// Mitsubishi GX Works2 project: B_v6_ladder   PLC: Q03UDE

PROGRAM MAIN
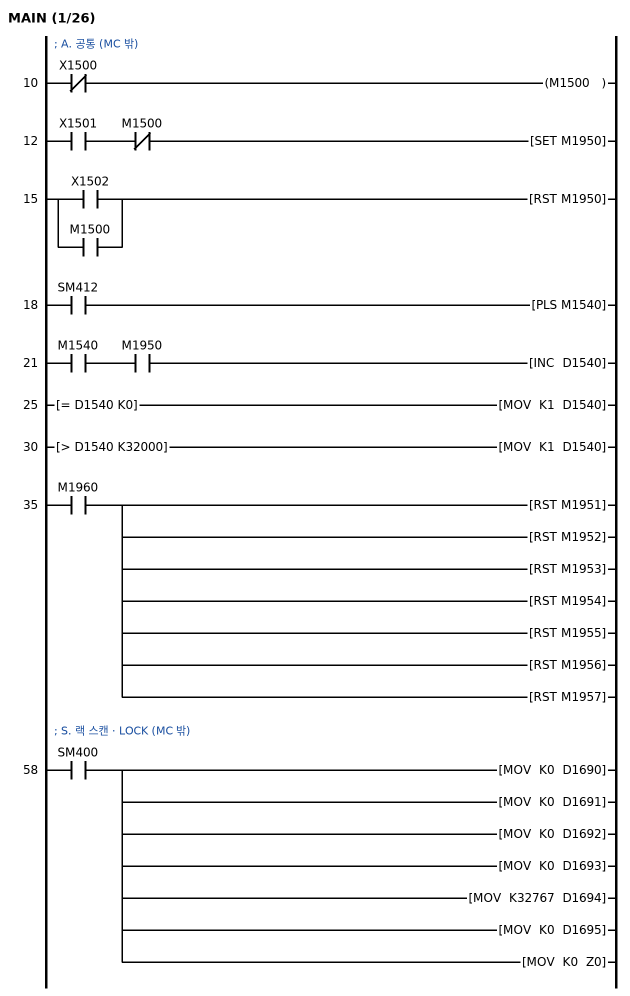
; A. 공통 (MC 밖)
10    LDI     X1500
      OUT     M1500
12    LD      X1501
      ANI     M1500
      SET     M1950
15    LD      X1502
      OR      M1500
      RST     M1950
18    LD      SM412
      PLS     M1540
21    LD      M1540
      AND     M1950
      INC     D1540
25    LD=     D1540 K0
      MOV     K1 D1540
30    LD>     D1540 K32000
      MOV     K1 D1540
35    LD      M1960
      RST     M1951
      RST     M1952
      RST     M1953
      RST     M1954
      RST     M1955
      RST     M1956
      RST     M1957
; S. 랙 스캔 · LOCK (MC 밖)
58    LD      SM400
      MOV     K0 D1690
      MOV     K0 D1691
      MOV     K0 D1692
      MOV     K0 D1693
      MOV     K32767 D1694
      MOV     K0 D1695
      MOV     K0 Z0
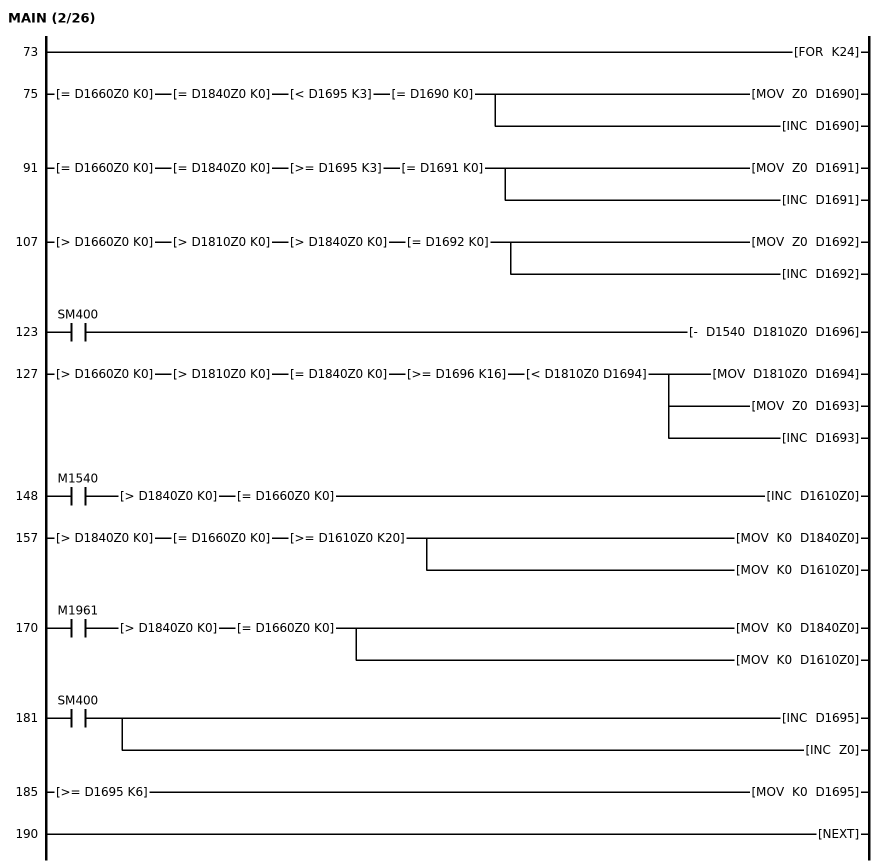
73    FOR     K24
75    LD=     D1660Z0 K0
      AND=    D1840Z0 K0
      AND<    D1695 K3
      AND=    D1690 K0
      MOV     Z0 D1690
      INC     D1690
91    LD=     D1660Z0 K0
      AND=    D1840Z0 K0
      AND>=   D1695 K3
      AND=    D1691 K0
      MOV     Z0 D1691
      INC     D1691
107   LD>     D1660Z0 K0
      AND>    D1810Z0 K0
      AND>    D1840Z0 K0
      AND=    D1692 K0
      MOV     Z0 D1692
      INC     D1692
123   LD      SM400
      -       D1540 D1810Z0 D1696
127   LD>     D1660Z0 K0
      AND>    D1810Z0 K0
      AND=    D1840Z0 K0
      AND>=   D1696 K16
      AND<    D1810Z0 D1694
      MOV     D1810Z0 D1694
      MOV     Z0 D1693
      INC     D1693
148   LD      M1540
      AND>    D1840Z0 K0
      AND=    D1660Z0 K0
      INC     D1610Z0
157   LD>     D1840Z0 K0
      AND=    D1660Z0 K0
      AND>=   D1610Z0 K20
      MOV     K0 D1840Z0
      MOV     K0 D1610Z0
170   LD      M1961
      AND>    D1840Z0 K0
      AND=    D1660Z0 K0
      MOV     K0 D1840Z0
      MOV     K0 D1610Z0
181   LD      SM400
      INC     D1695
      INC     Z0
185   LD>=    D1695 K6
      MOV     K0 D1695
190   NEXT
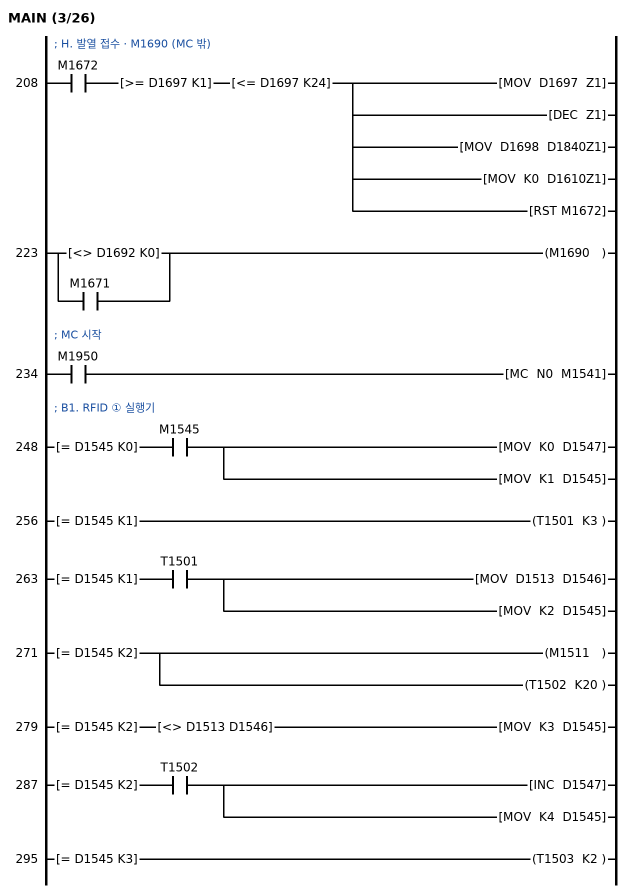
; H. 발열 접수 · M1690 (MC 밖)
208   LD      M1672
      AND>=   D1697 K1
      AND<=   D1697 K24
      MOV     D1697 Z1
      DEC     Z1
      MOV     D1698 D1840Z1
      MOV     K0 D1610Z1
      RST     M1672
223   LD<>    D1692 K0
      OR      M1671
      OUT     M1690
; MC 시작
234   LD      M1950
      MC      N0 M1541
; B1. RFID ① 실행기
248   LD=     D1545 K0
      AND     M1545
      MOV     K0 D1547
      MOV     K1 D1545
256   LD=     D1545 K1
      OUT     T1501 K3
263   LD=     D1545 K1
      AND     T1501
      MOV     D1513 D1546
      MOV     K2 D1545
271   LD=     D1545 K2
      OUT     M1511
      OUT     T1502 K20
279   LD=     D1545 K2
      AND<>   D1513 D1546
      MOV     K3 D1545
287   LD=     D1545 K2
      AND     T1502
      INC     D1547
      MOV     K4 D1545
295   LD=     D1545 K3
      OUT     T1503 K2
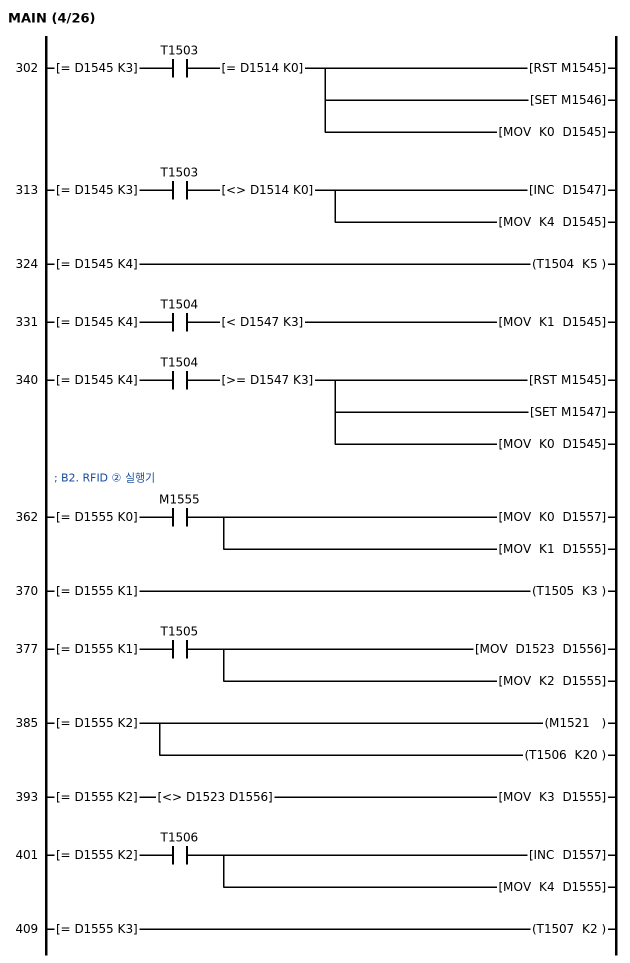
302   LD=     D1545 K3
      AND     T1503
      AND=    D1514 K0
      RST     M1545
      SET     M1546
      MOV     K0 D1545
313   LD=     D1545 K3
      AND     T1503
      AND<>   D1514 K0
      INC     D1547
      MOV     K4 D1545
324   LD=     D1545 K4
      OUT     T1504 K5
331   LD=     D1545 K4
      AND     T1504
      AND<    D1547 K3
      MOV     K1 D1545
340   LD=     D1545 K4
      AND     T1504
      AND>=   D1547 K3
      RST     M1545
      SET     M1547
      MOV     K0 D1545
; B2. RFID ② 실행기
362   LD=     D1555 K0
      AND     M1555
      MOV     K0 D1557
      MOV     K1 D1555
370   LD=     D1555 K1
      OUT     T1505 K3
377   LD=     D1555 K1
      AND     T1505
      MOV     D1523 D1556
      MOV     K2 D1555
385   LD=     D1555 K2
      OUT     M1521
      OUT     T1506 K20
393   LD=     D1555 K2
      AND<>   D1523 D1556
      MOV     K3 D1555
401   LD=     D1555 K2
      AND     T1506
      INC     D1557
      MOV     K4 D1555
409   LD=     D1555 K3
      OUT     T1507 K2
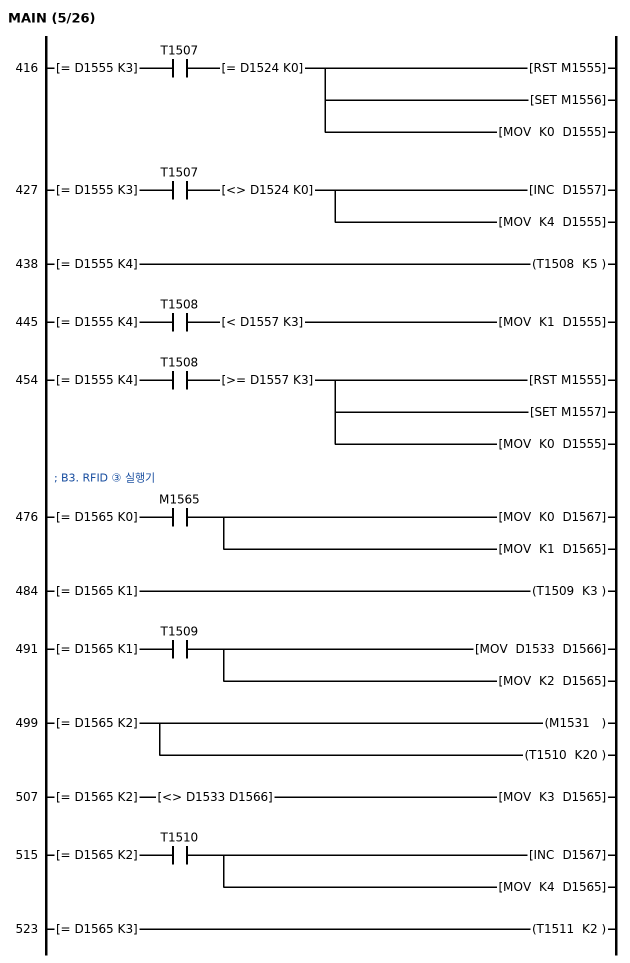
416   LD=     D1555 K3
      AND     T1507
      AND=    D1524 K0
      RST     M1555
      SET     M1556
      MOV     K0 D1555
427   LD=     D1555 K3
      AND     T1507
      AND<>   D1524 K0
      INC     D1557
      MOV     K4 D1555
438   LD=     D1555 K4
      OUT     T1508 K5
445   LD=     D1555 K4
      AND     T1508
      AND<    D1557 K3
      MOV     K1 D1555
454   LD=     D1555 K4
      AND     T1508
      AND>=   D1557 K3
      RST     M1555
      SET     M1557
      MOV     K0 D1555
; B3. RFID ③ 실행기
476   LD=     D1565 K0
      AND     M1565
      MOV     K0 D1567
      MOV     K1 D1565
484   LD=     D1565 K1
      OUT     T1509 K3
491   LD=     D1565 K1
      AND     T1509
      MOV     D1533 D1566
      MOV     K2 D1565
499   LD=     D1565 K2
      OUT     M1531
      OUT     T1510 K20
507   LD=     D1565 K2
      AND<>   D1533 D1566
      MOV     K3 D1565
515   LD=     D1565 K2
      AND     T1510
      INC     D1567
      MOV     K4 D1565
523   LD=     D1565 K3
      OUT     T1511 K2
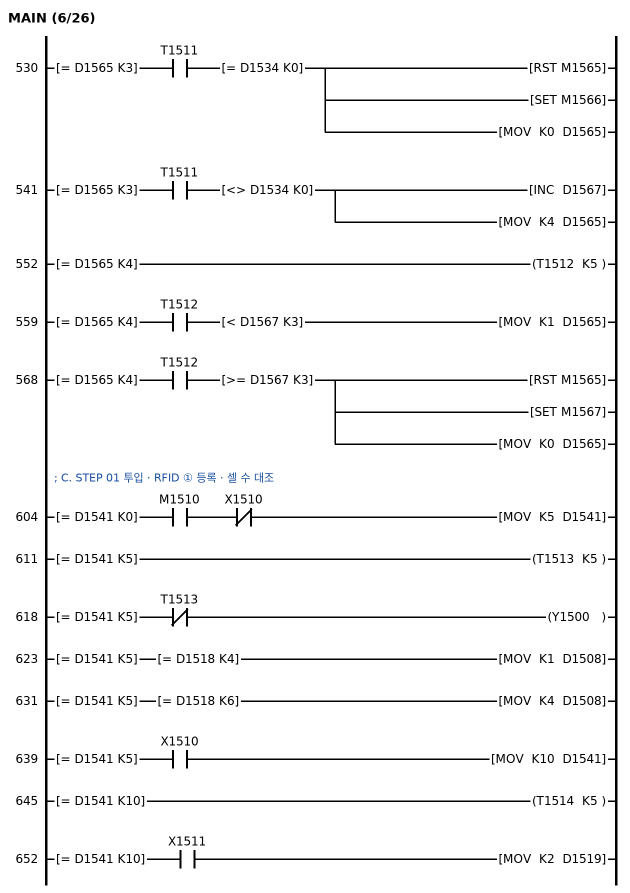
530   LD=     D1565 K3
      AND     T1511
      AND=    D1534 K0
      RST     M1565
      SET     M1566
      MOV     K0 D1565
541   LD=     D1565 K3
      AND     T1511
      AND<>   D1534 K0
      INC     D1567
      MOV     K4 D1565
552   LD=     D1565 K4
      OUT     T1512 K5
559   LD=     D1565 K4
      AND     T1512
      AND<    D1567 K3
      MOV     K1 D1565
568   LD=     D1565 K4
      AND     T1512
      AND>=   D1567 K3
      RST     M1565
      SET     M1567
      MOV     K0 D1565
; C. STEP 01 투입 · RFID ① 등록 · 셀 수 대조
604   LD=     D1541 K0
      AND     M1510
      ANI     X1510
      MOV     K5 D1541
611   LD=     D1541 K5
      OUT     T1513 K5
618   LD=     D1541 K5
      ANI     T1513
      OUT     Y1500
623   LD=     D1541 K5
      AND=    D1518 K4
      MOV     K1 D1508
631   LD=     D1541 K5
      AND=    D1518 K6
      MOV     K4 D1508
639   LD=     D1541 K5
      AND     X1510
      MOV     K10 D1541
645   LD=     D1541 K10
      OUT     T1514 K5
652   LD=     D1541 K10
      AND     X1511
      MOV     K2 D1519
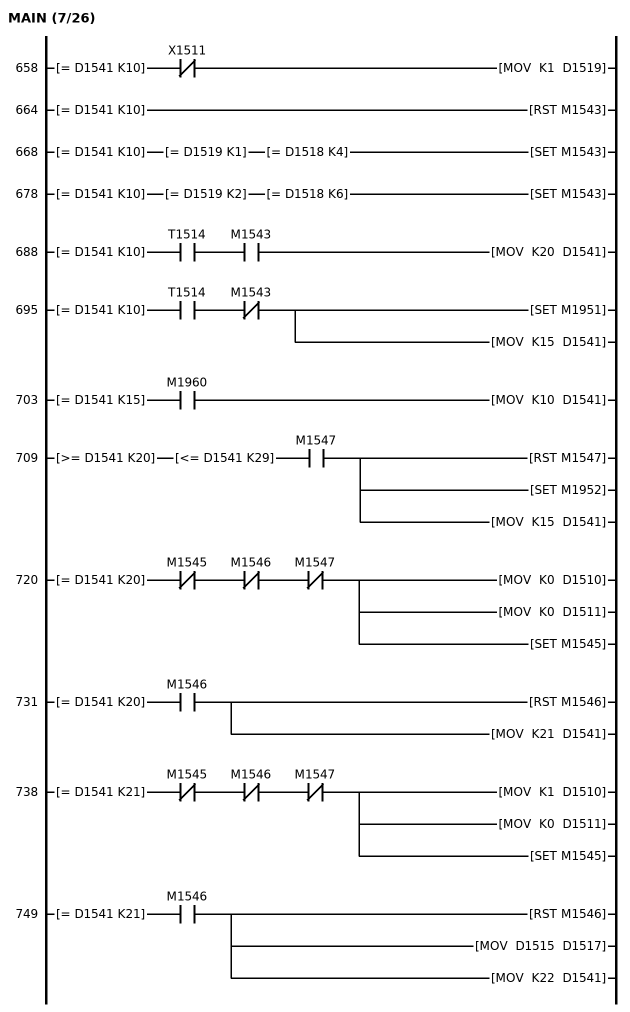
658   LD=     D1541 K10
      ANI     X1511
      MOV     K1 D1519
664   LD=     D1541 K10
      RST     M1543
668   LD=     D1541 K10
      AND=    D1519 K1
      AND=    D1518 K4
      SET     M1543
678   LD=     D1541 K10
      AND=    D1519 K2
      AND=    D1518 K6
      SET     M1543
688   LD=     D1541 K10
      AND     T1514
      AND     M1543
      MOV     K20 D1541
695   LD=     D1541 K10
      AND     T1514
      ANI     M1543
      SET     M1951
      MOV     K15 D1541
703   LD=     D1541 K15
      AND     M1960
      MOV     K10 D1541
709   LD>=    D1541 K20
      AND<=   D1541 K29
      AND     M1547
      RST     M1547
      SET     M1952
      MOV     K15 D1541
720   LD=     D1541 K20
      ANI     M1545
      ANI     M1546
      ANI     M1547
      MOV     K0 D1510
      MOV     K0 D1511
      SET     M1545
731   LD=     D1541 K20
      AND     M1546
      RST     M1546
      MOV     K21 D1541
738   LD=     D1541 K21
      ANI     M1545
      ANI     M1546
      ANI     M1547
      MOV     K1 D1510
      MOV     K0 D1511
      SET     M1545
749   LD=     D1541 K21
      AND     M1546
      RST     M1546
      MOV     D1515 D1517
      MOV     K22 D1541
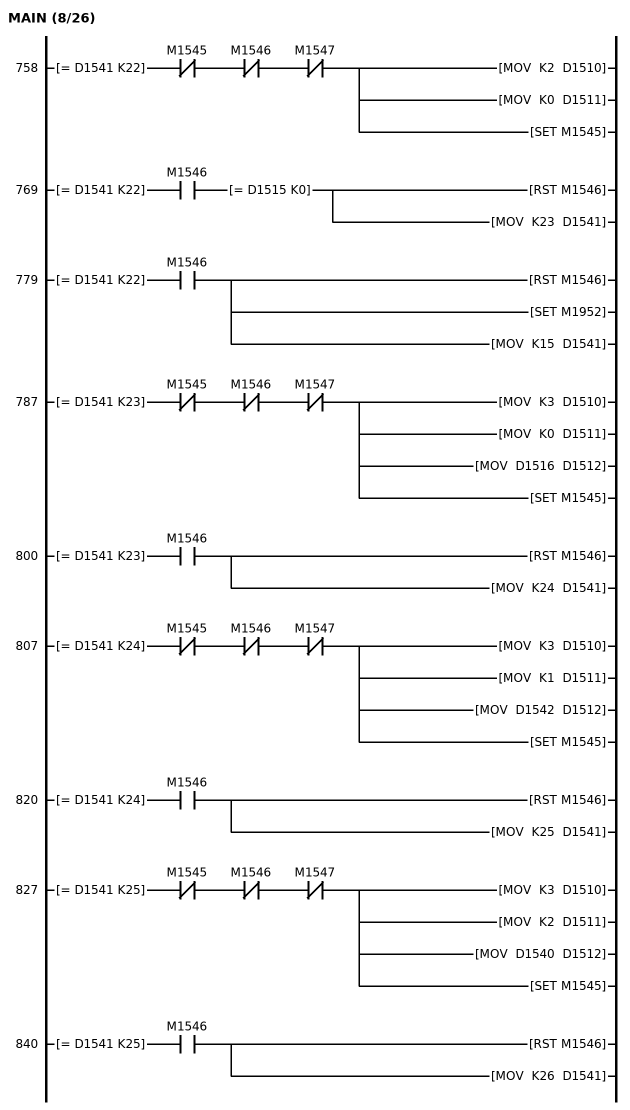
758   LD=     D1541 K22
      ANI     M1545
      ANI     M1546
      ANI     M1547
      MOV     K2 D1510
      MOV     K0 D1511
      SET     M1545
769   LD=     D1541 K22
      AND     M1546
      AND=    D1515 K0
      RST     M1546
      MOV     K23 D1541
779   LD=     D1541 K22
      AND     M1546
      RST     M1546
      SET     M1952
      MOV     K15 D1541
787   LD=     D1541 K23
      ANI     M1545
      ANI     M1546
      ANI     M1547
      MOV     K3 D1510
      MOV     K0 D1511
      MOV     D1516 D1512
      SET     M1545
800   LD=     D1541 K23
      AND     M1546
      RST     M1546
      MOV     K24 D1541
807   LD=     D1541 K24
      ANI     M1545
      ANI     M1546
      ANI     M1547
      MOV     K3 D1510
      MOV     K1 D1511
      MOV     D1542 D1512
      SET     M1545
820   LD=     D1541 K24
      AND     M1546
      RST     M1546
      MOV     K25 D1541
827   LD=     D1541 K25
      ANI     M1545
      ANI     M1546
      ANI     M1547
      MOV     K3 D1510
      MOV     K2 D1511
      MOV     D1540 D1512
      SET     M1545
840   LD=     D1541 K25
      AND     M1546
      RST     M1546
      MOV     K26 D1541
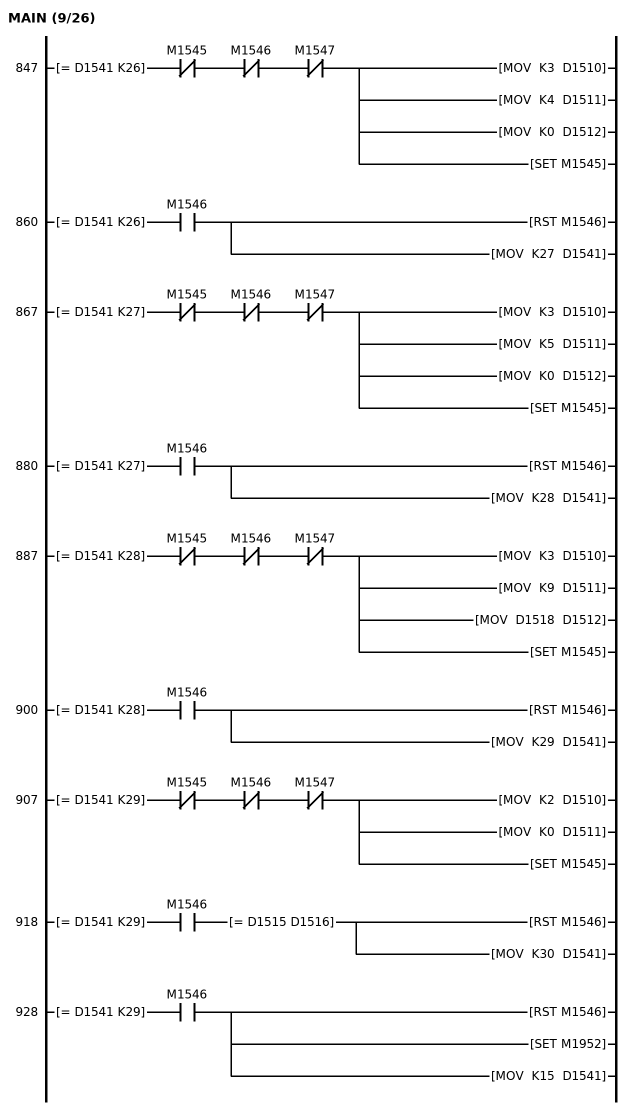
847   LD=     D1541 K26
      ANI     M1545
      ANI     M1546
      ANI     M1547
      MOV     K3 D1510
      MOV     K4 D1511
      MOV     K0 D1512
      SET     M1545
860   LD=     D1541 K26
      AND     M1546
      RST     M1546
      MOV     K27 D1541
867   LD=     D1541 K27
      ANI     M1545
      ANI     M1546
      ANI     M1547
      MOV     K3 D1510
      MOV     K5 D1511
      MOV     K0 D1512
      SET     M1545
880   LD=     D1541 K27
      AND     M1546
      RST     M1546
      MOV     K28 D1541
887   LD=     D1541 K28
      ANI     M1545
      ANI     M1546
      ANI     M1547
      MOV     K3 D1510
      MOV     K9 D1511
      MOV     D1518 D1512
      SET     M1545
900   LD=     D1541 K28
      AND     M1546
      RST     M1546
      MOV     K29 D1541
907   LD=     D1541 K29
      ANI     M1545
      ANI     M1546
      ANI     M1547
      MOV     K2 D1510
      MOV     K0 D1511
      SET     M1545
918   LD=     D1541 K29
      AND     M1546
      AND=    D1515 D1516
      RST     M1546
      MOV     K30 D1541
928   LD=     D1541 K29
      AND     M1546
      RST     M1546
      SET     M1952
      MOV     K15 D1541
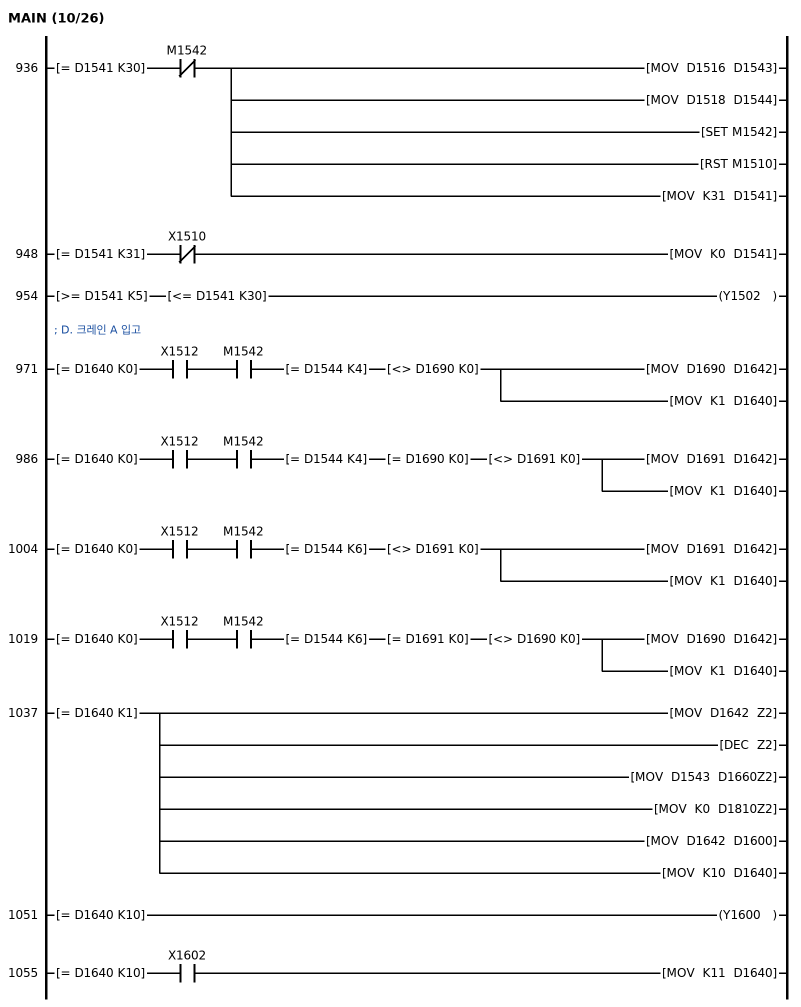
936   LD=     D1541 K30
      ANI     M1542
      MOV     D1516 D1543
      MOV     D1518 D1544
      SET     M1542
      RST     M1510
      MOV     K31 D1541
948   LD=     D1541 K31
      ANI     X1510
      MOV     K0 D1541
954   LD>=    D1541 K5
      AND<=   D1541 K30
      OUT     Y1502
; D. 크레인 A 입고
971   LD=     D1640 K0
      AND     X1512
      AND     M1542
      AND=    D1544 K4
      AND<>   D1690 K0
      MOV     D1690 D1642
      MOV     K1 D1640
986   LD=     D1640 K0
      AND     X1512
      AND     M1542
      AND=    D1544 K4
      AND=    D1690 K0
      AND<>   D1691 K0
      MOV     D1691 D1642
      MOV     K1 D1640
1004  LD=     D1640 K0
      AND     X1512
      AND     M1542
      AND=    D1544 K6
      AND<>   D1691 K0
      MOV     D1691 D1642
      MOV     K1 D1640
1019  LD=     D1640 K0
      AND     X1512
      AND     M1542
      AND=    D1544 K6
      AND=    D1691 K0
      AND<>   D1690 K0
      MOV     D1690 D1642
      MOV     K1 D1640
1037  LD=     D1640 K1
      MOV     D1642 Z2
      DEC     Z2
      MOV     D1543 D1660Z2
      MOV     K0 D1810Z2
      MOV     D1642 D1600
      MOV     K10 D1640
1051  LD=     D1640 K10
      OUT     Y1600
1055  LD=     D1640 K10
      AND     X1602
      MOV     K11 D1640
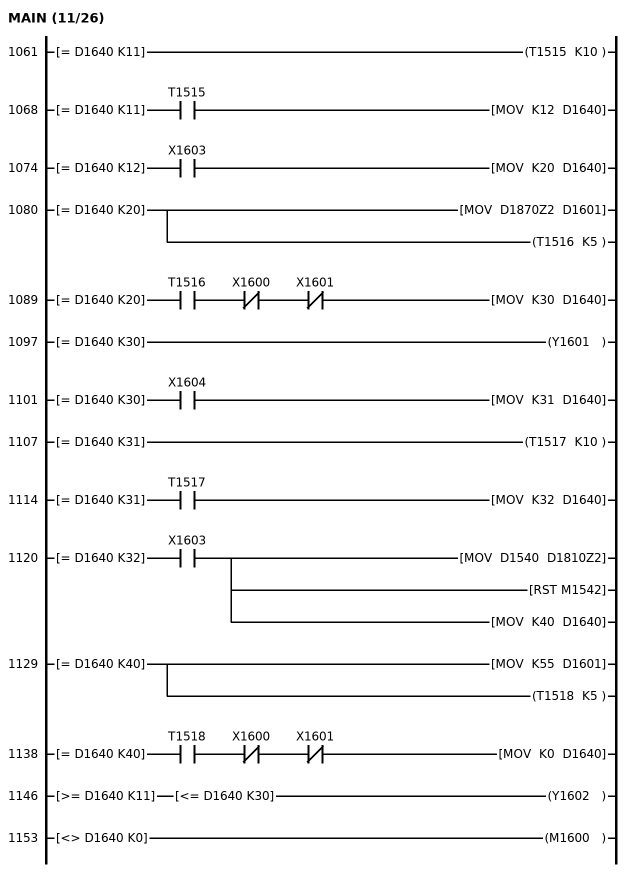
1061  LD=     D1640 K11
      OUT     T1515 K10
1068  LD=     D1640 K11
      AND     T1515
      MOV     K12 D1640
1074  LD=     D1640 K12
      AND     X1603
      MOV     K20 D1640
1080  LD=     D1640 K20
      MOV     D1870Z2 D1601
      OUT     T1516 K5
1089  LD=     D1640 K20
      AND     T1516
      ANI     X1600
      ANI     X1601
      MOV     K30 D1640
1097  LD=     D1640 K30
      OUT     Y1601
1101  LD=     D1640 K30
      AND     X1604
      MOV     K31 D1640
1107  LD=     D1640 K31
      OUT     T1517 K10
1114  LD=     D1640 K31
      AND     T1517
      MOV     K32 D1640
1120  LD=     D1640 K32
      AND     X1603
      MOV     D1540 D1810Z2
      RST     M1542
      MOV     K40 D1640
1129  LD=     D1640 K40
      MOV     K55 D1601
      OUT     T1518 K5
1138  LD=     D1640 K40
      AND     T1518
      ANI     X1600
      ANI     X1601
      MOV     K0 D1640
1146  LD>=    D1640 K11
      AND<=   D1640 K30
      OUT     Y1602
1153  LD<>    D1640 K0
      OUT     M1600
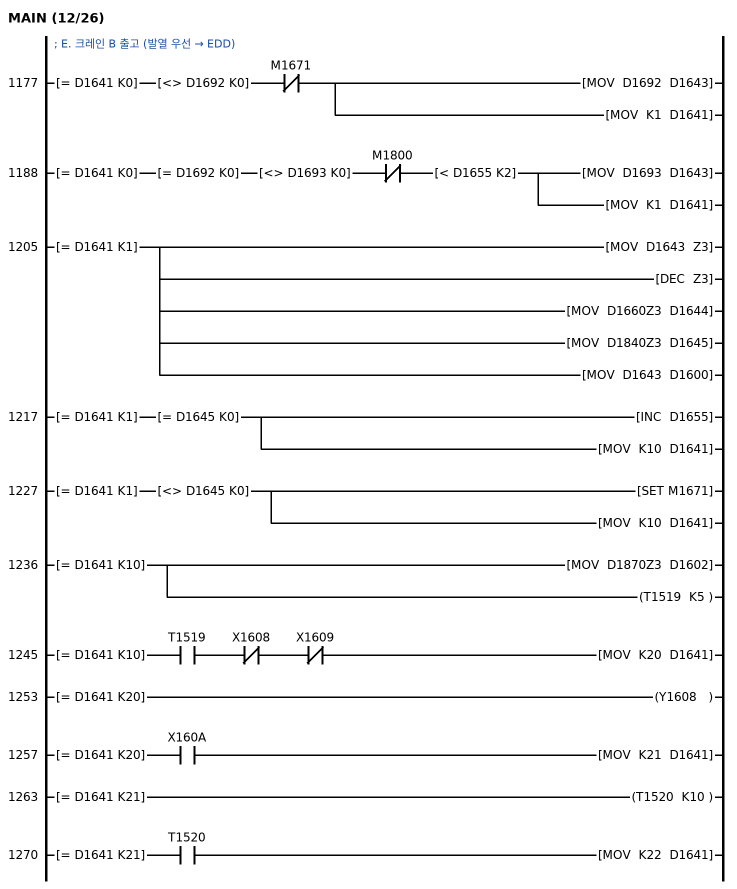
; E. 크레인 B 출고 (발열 우선 → EDD)
1177  LD=     D1641 K0
      AND<>   D1692 K0
      ANI     M1671
      MOV     D1692 D1643
      MOV     K1 D1641
1188  LD=     D1641 K0
      AND=    D1692 K0
      AND<>   D1693 K0
      ANI     M1800
      AND<    D1655 K2
      MOV     D1693 D1643
      MOV     K1 D1641
1205  LD=     D1641 K1
      MOV     D1643 Z3
      DEC     Z3
      MOV     D1660Z3 D1644
      MOV     D1840Z3 D1645
      MOV     D1643 D1600
1217  LD=     D1641 K1
      AND=    D1645 K0
      INC     D1655
      MOV     K10 D1641
1227  LD=     D1641 K1
      AND<>   D1645 K0
      SET     M1671
      MOV     K10 D1641
1236  LD=     D1641 K10
      MOV     D1870Z3 D1602
      OUT     T1519 K5
1245  LD=     D1641 K10
      AND     T1519
      ANI     X1608
      ANI     X1609
      MOV     K20 D1641
1253  LD=     D1641 K20
      OUT     Y1608
1257  LD=     D1641 K20
      AND     X160A
      MOV     K21 D1641
1263  LD=     D1641 K21
      OUT     T1520 K10
1270  LD=     D1641 K21
      AND     T1520
      MOV     K22 D1641
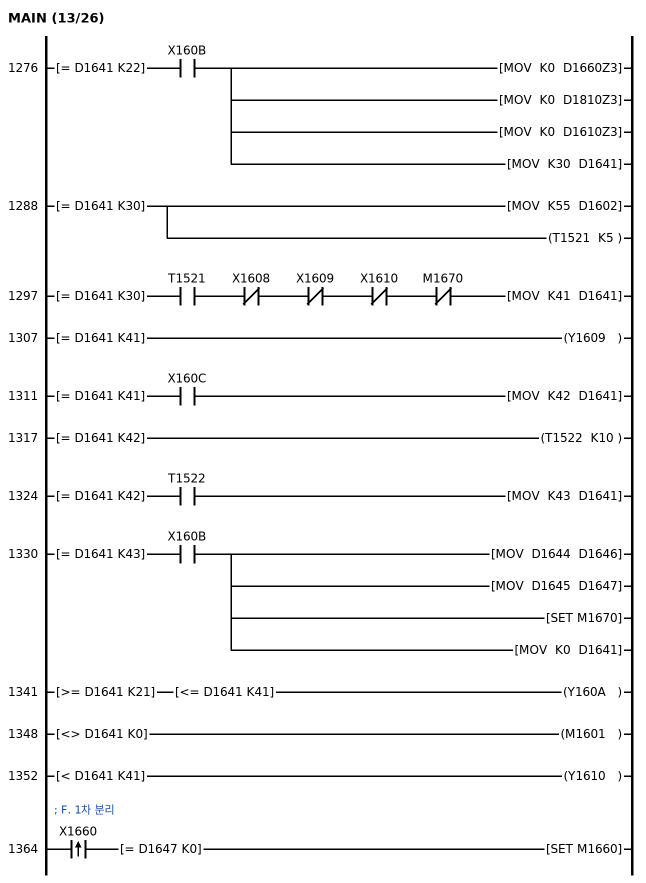
1276  LD=     D1641 K22
      AND     X160B
      MOV     K0 D1660Z3
      MOV     K0 D1810Z3
      MOV     K0 D1610Z3
      MOV     K30 D1641
1288  LD=     D1641 K30
      MOV     K55 D1602
      OUT     T1521 K5
1297  LD=     D1641 K30
      AND     T1521
      ANI     X1608
      ANI     X1609
      ANI     X1610
      ANI     M1670
      MOV     K41 D1641
1307  LD=     D1641 K41
      OUT     Y1609
1311  LD=     D1641 K41
      AND     X160C
      MOV     K42 D1641
1317  LD=     D1641 K42
      OUT     T1522 K10
1324  LD=     D1641 K42
      AND     T1522
      MOV     K43 D1641
1330  LD=     D1641 K43
      AND     X160B
      MOV     D1644 D1646
      MOV     D1645 D1647
      SET     M1670
      MOV     K0 D1641
1341  LD>=    D1641 K21
      AND<=   D1641 K41
      OUT     Y160A
1348  LD<>    D1641 K0
      OUT     M1601
1352  LD<     D1641 K41
      OUT     Y1610
; F. 1차 분리
1364  LDP     X1660
      AND=    D1647 K0
      SET     M1660
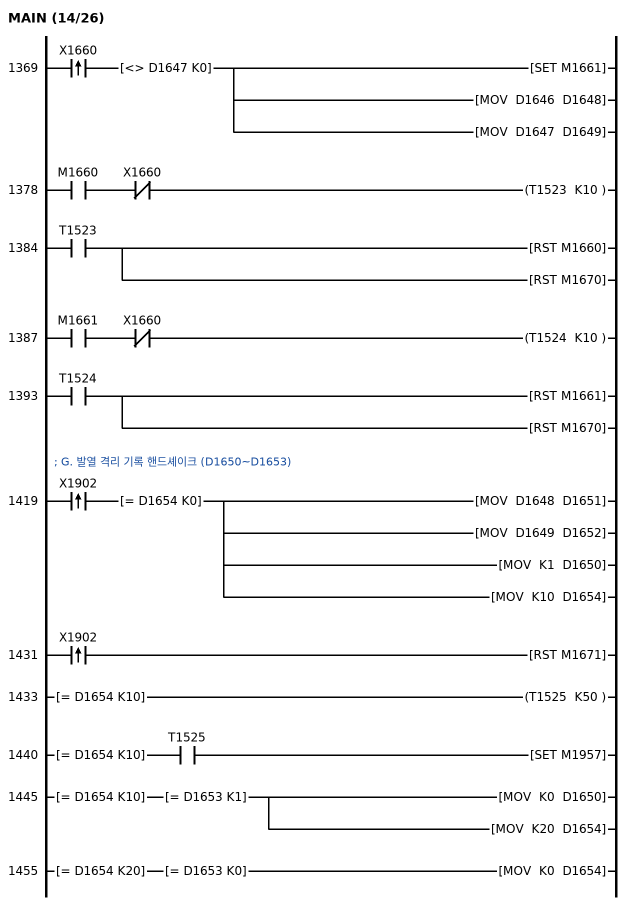
1369  LDP     X1660
      AND<>   D1647 K0
      SET     M1661
      MOV     D1646 D1648
      MOV     D1647 D1649
1378  LD      M1660
      ANI     X1660
      OUT     T1523 K10
1384  LD      T1523
      RST     M1660
      RST     M1670
1387  LD      M1661
      ANI     X1660
      OUT     T1524 K10
1393  LD      T1524
      RST     M1661
      RST     M1670
; G. 발열 격리 기록 핸드셰이크 (D1650~D1653)
1419  LDP     X1902
      AND=    D1654 K0
      MOV     D1648 D1651
      MOV     D1649 D1652
      MOV     K1 D1650
      MOV     K10 D1654
1431  LDP     X1902
      RST     M1671
1433  LD=     D1654 K10
      OUT     T1525 K50
1440  LD=     D1654 K10
      AND     T1525
      SET     M1957
1445  LD=     D1654 K10
      AND=    D1653 K1
      MOV     K0 D1650
      MOV     K20 D1654
1455  LD=     D1654 K20
      AND=    D1653 K0
      MOV     K0 D1654
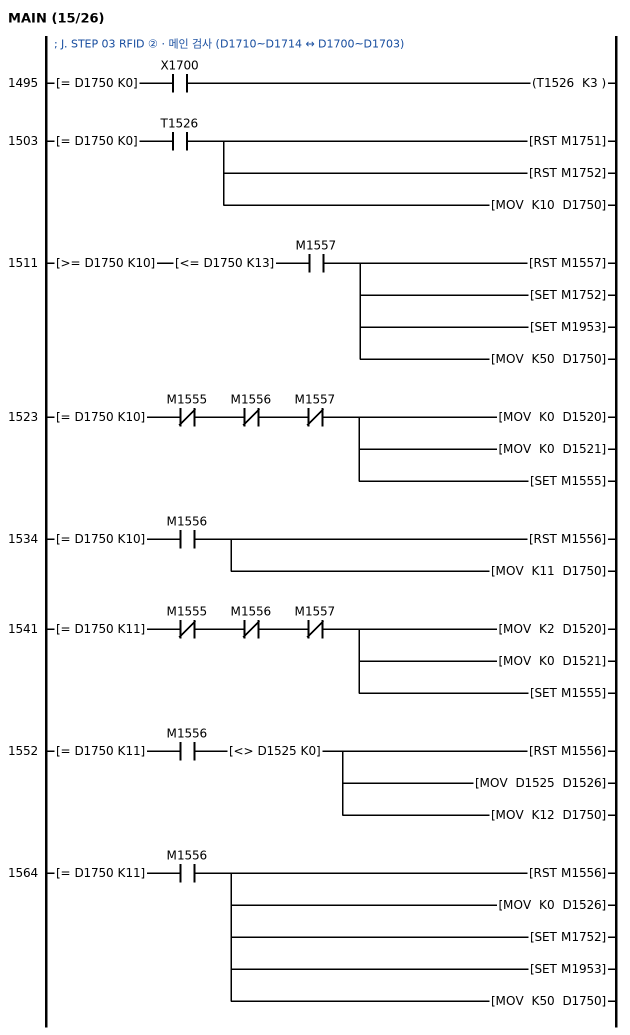
; J. STEP 03 RFID ② · 메인 검사 (D1710~D1714 ↔ D1700~D1703)
1495  LD=     D1750 K0
      AND     X1700
      OUT     T1526 K3
1503  LD=     D1750 K0
      AND     T1526
      RST     M1751
      RST     M1752
      MOV     K10 D1750
1511  LD>=    D1750 K10
      AND<=   D1750 K13
      AND     M1557
      RST     M1557
      SET     M1752
      SET     M1953
      MOV     K50 D1750
1523  LD=     D1750 K10
      ANI     M1555
      ANI     M1556
      ANI     M1557
      MOV     K0 D1520
      MOV     K0 D1521
      SET     M1555
1534  LD=     D1750 K10
      AND     M1556
      RST     M1556
      MOV     K11 D1750
1541  LD=     D1750 K11
      ANI     M1555
      ANI     M1556
      ANI     M1557
      MOV     K2 D1520
      MOV     K0 D1521
      SET     M1555
1552  LD=     D1750 K11
      AND     M1556
      AND<>   D1525 K0
      RST     M1556
      MOV     D1525 D1526
      MOV     K12 D1750
1564  LD=     D1750 K11
      AND     M1556
      RST     M1556
      MOV     K0 D1526
      SET     M1752
      SET     M1953
      MOV     K50 D1750
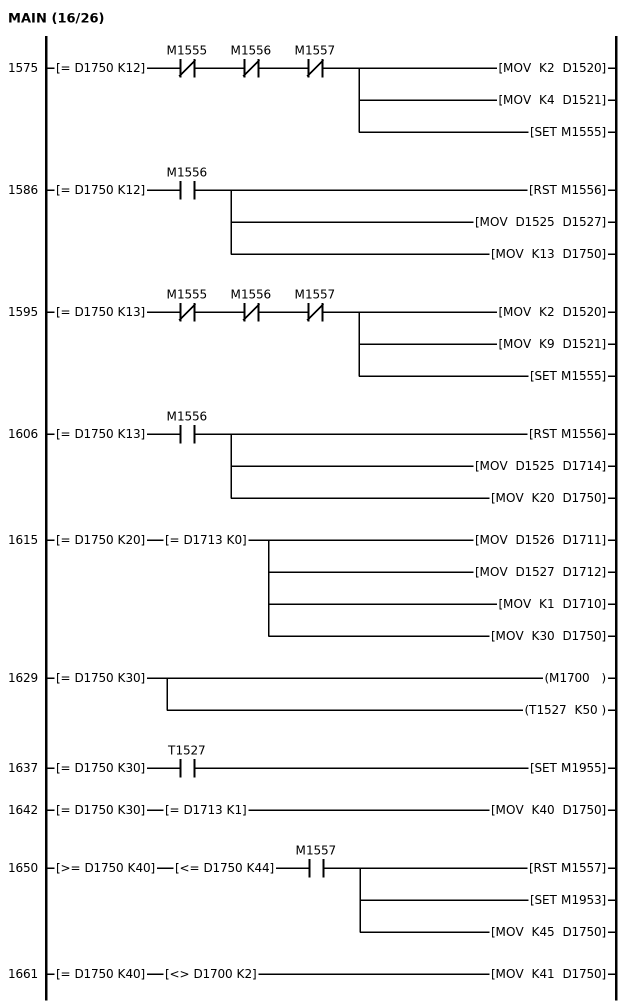
1575  LD=     D1750 K12
      ANI     M1555
      ANI     M1556
      ANI     M1557
      MOV     K2 D1520
      MOV     K4 D1521
      SET     M1555
1586  LD=     D1750 K12
      AND     M1556
      RST     M1556
      MOV     D1525 D1527
      MOV     K13 D1750
1595  LD=     D1750 K13
      ANI     M1555
      ANI     M1556
      ANI     M1557
      MOV     K2 D1520
      MOV     K9 D1521
      SET     M1555
1606  LD=     D1750 K13
      AND     M1556
      RST     M1556
      MOV     D1525 D1714
      MOV     K20 D1750
1615  LD=     D1750 K20
      AND=    D1713 K0
      MOV     D1526 D1711
      MOV     D1527 D1712
      MOV     K1 D1710
      MOV     K30 D1750
1629  LD=     D1750 K30
      OUT     M1700
      OUT     T1527 K50
1637  LD=     D1750 K30
      AND     T1527
      SET     M1955
1642  LD=     D1750 K30
      AND=    D1713 K1
      MOV     K40 D1750
1650  LD>=    D1750 K40
      AND<=   D1750 K44
      AND     M1557
      RST     M1557
      SET     M1953
      MOV     K45 D1750
1661  LD=     D1750 K40
      AND<>   D1700 K2
      MOV     K41 D1750
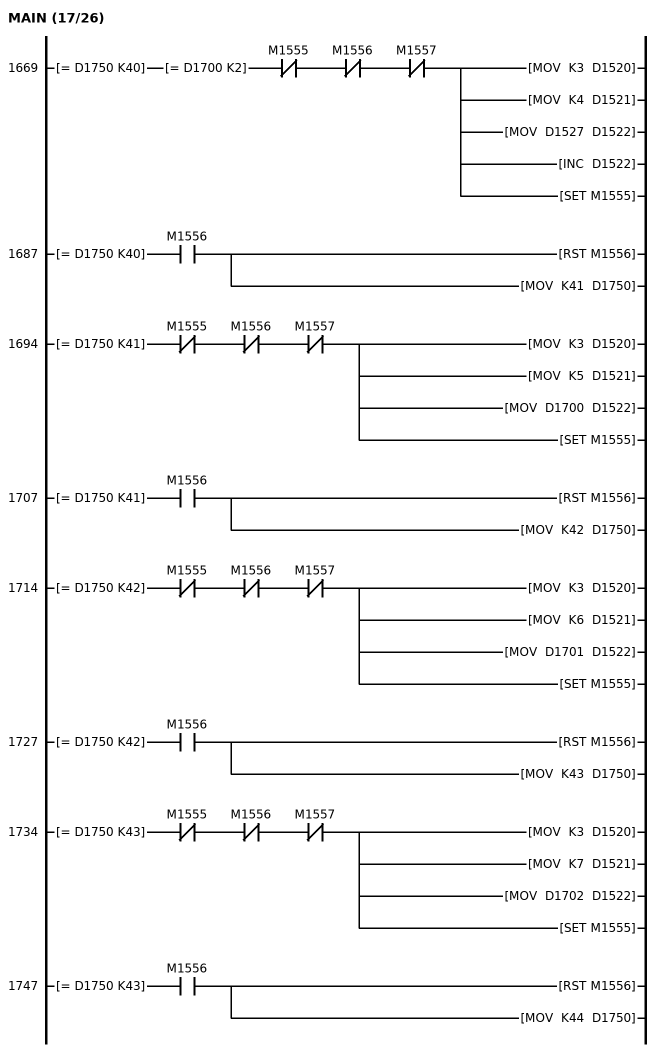
1669  LD=     D1750 K40
      AND=    D1700 K2
      ANI     M1555
      ANI     M1556
      ANI     M1557
      MOV     K3 D1520
      MOV     K4 D1521
      MOV     D1527 D1522
      INC     D1522
      SET     M1555
1687  LD=     D1750 K40
      AND     M1556
      RST     M1556
      MOV     K41 D1750
1694  LD=     D1750 K41
      ANI     M1555
      ANI     M1556
      ANI     M1557
      MOV     K3 D1520
      MOV     K5 D1521
      MOV     D1700 D1522
      SET     M1555
1707  LD=     D1750 K41
      AND     M1556
      RST     M1556
      MOV     K42 D1750
1714  LD=     D1750 K42
      ANI     M1555
      ANI     M1556
      ANI     M1557
      MOV     K3 D1520
      MOV     K6 D1521
      MOV     D1701 D1522
      SET     M1555
1727  LD=     D1750 K42
      AND     M1556
      RST     M1556
      MOV     K43 D1750
1734  LD=     D1750 K43
      ANI     M1555
      ANI     M1556
      ANI     M1557
      MOV     K3 D1520
      MOV     K7 D1521
      MOV     D1702 D1522
      SET     M1555
1747  LD=     D1750 K43
      AND     M1556
      RST     M1556
      MOV     K44 D1750
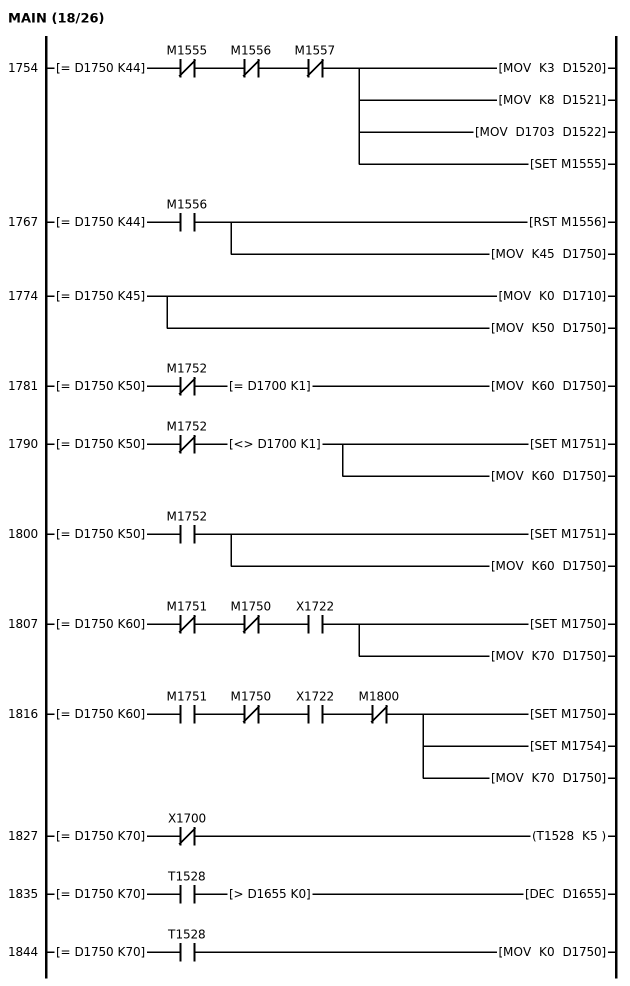
1754  LD=     D1750 K44
      ANI     M1555
      ANI     M1556
      ANI     M1557
      MOV     K3 D1520
      MOV     K8 D1521
      MOV     D1703 D1522
      SET     M1555
1767  LD=     D1750 K44
      AND     M1556
      RST     M1556
      MOV     K45 D1750
1774  LD=     D1750 K45
      MOV     K0 D1710
      MOV     K50 D1750
1781  LD=     D1750 K50
      ANI     M1752
      AND=    D1700 K1
      MOV     K60 D1750
1790  LD=     D1750 K50
      ANI     M1752
      AND<>   D1700 K1
      SET     M1751
      MOV     K60 D1750
1800  LD=     D1750 K50
      AND     M1752
      SET     M1751
      MOV     K60 D1750
1807  LD=     D1750 K60
      ANI     M1751
      ANI     M1750
      AND     X1722
      SET     M1750
      MOV     K70 D1750
1816  LD=     D1750 K60
      AND     M1751
      ANI     M1750
      AND     X1722
      ANI     M1800
      SET     M1750
      SET     M1754
      MOV     K70 D1750
1827  LD=     D1750 K70
      ANI     X1700
      OUT     T1528 K5
1835  LD=     D1750 K70
      AND     T1528
      AND>    D1655 K0
      DEC     D1655
1844  LD=     D1750 K70
      AND     T1528
      MOV     K0 D1750
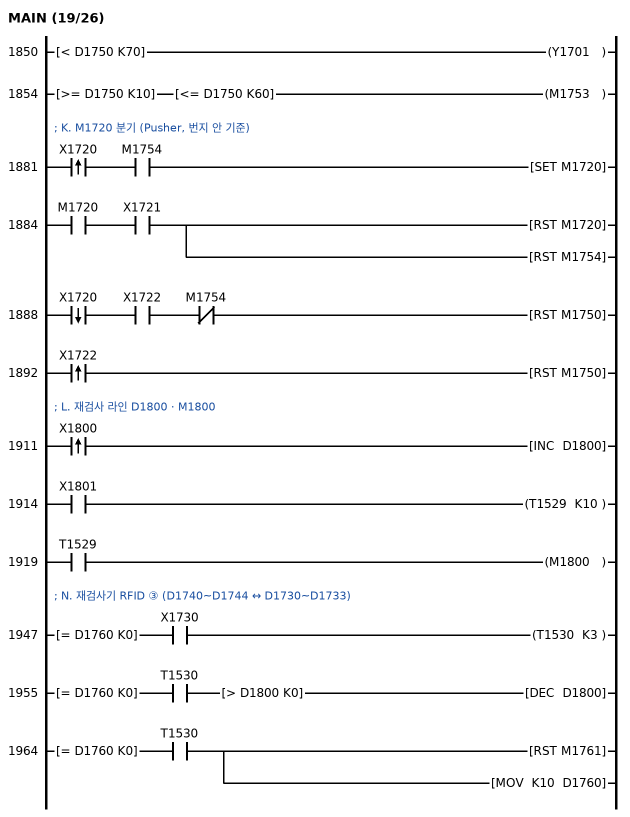
1850  LD<     D1750 K70
      OUT     Y1701
1854  LD>=    D1750 K10
      AND<=   D1750 K60
      OUT     M1753
; K. M1720 분기 (Pusher, 번지 안 기준)
1881  LDP     X1720
      AND     M1754
      SET     M1720
1884  LD      M1720
      AND     X1721
      RST     M1720
      RST     M1754
1888  LDF     X1720
      AND     X1722
      ANI     M1754
      RST     M1750
1892  LDP     X1722
      RST     M1750
; L. 재검사 라인 D1800 · M1800
1911  LDP     X1800
      INC     D1800
1914  LD      X1801
      OUT     T1529 K10
1919  LD      T1529
      OUT     M1800
; N. 재검사기 RFID ③ (D1740~D1744 ↔ D1730~D1733)
1947  LD=     D1760 K0
      AND     X1730
      OUT     T1530 K3
1955  LD=     D1760 K0
      AND     T1530
      AND>    D1800 K0
      DEC     D1800
1964  LD=     D1760 K0
      AND     T1530
      RST     M1761
      MOV     K10 D1760
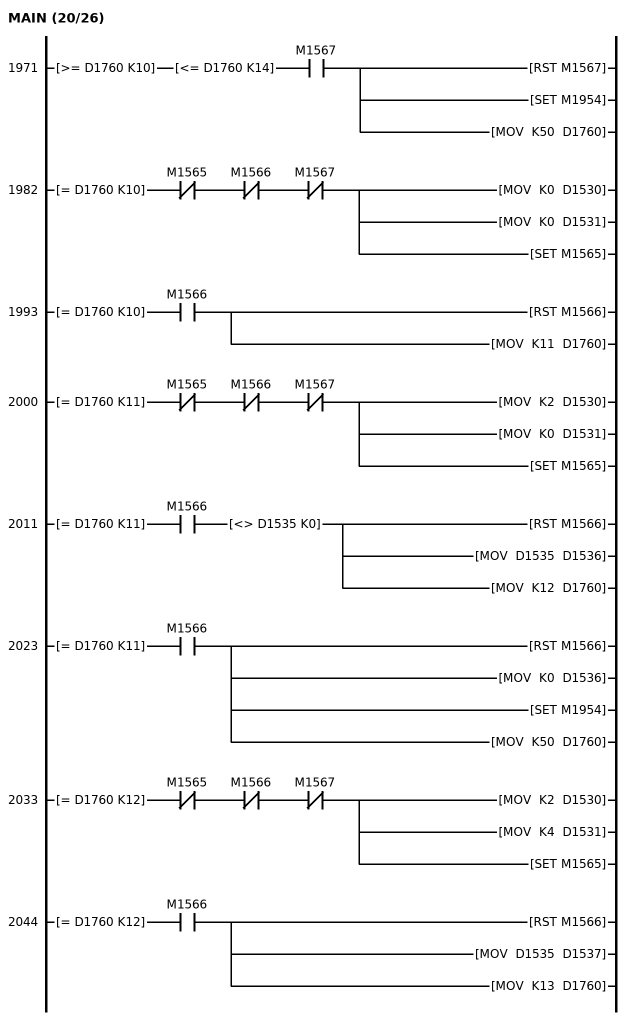
1971  LD>=    D1760 K10
      AND<=   D1760 K14
      AND     M1567
      RST     M1567
      SET     M1954
      MOV     K50 D1760
1982  LD=     D1760 K10
      ANI     M1565
      ANI     M1566
      ANI     M1567
      MOV     K0 D1530
      MOV     K0 D1531
      SET     M1565
1993  LD=     D1760 K10
      AND     M1566
      RST     M1566
      MOV     K11 D1760
2000  LD=     D1760 K11
      ANI     M1565
      ANI     M1566
      ANI     M1567
      MOV     K2 D1530
      MOV     K0 D1531
      SET     M1565
2011  LD=     D1760 K11
      AND     M1566
      AND<>   D1535 K0
      RST     M1566
      MOV     D1535 D1536
      MOV     K12 D1760
2023  LD=     D1760 K11
      AND     M1566
      RST     M1566
      MOV     K0 D1536
      SET     M1954
      MOV     K50 D1760
2033  LD=     D1760 K12
      ANI     M1565
      ANI     M1566
      ANI     M1567
      MOV     K2 D1530
      MOV     K4 D1531
      SET     M1565
2044  LD=     D1760 K12
      AND     M1566
      RST     M1566
      MOV     D1535 D1537
      MOV     K13 D1760
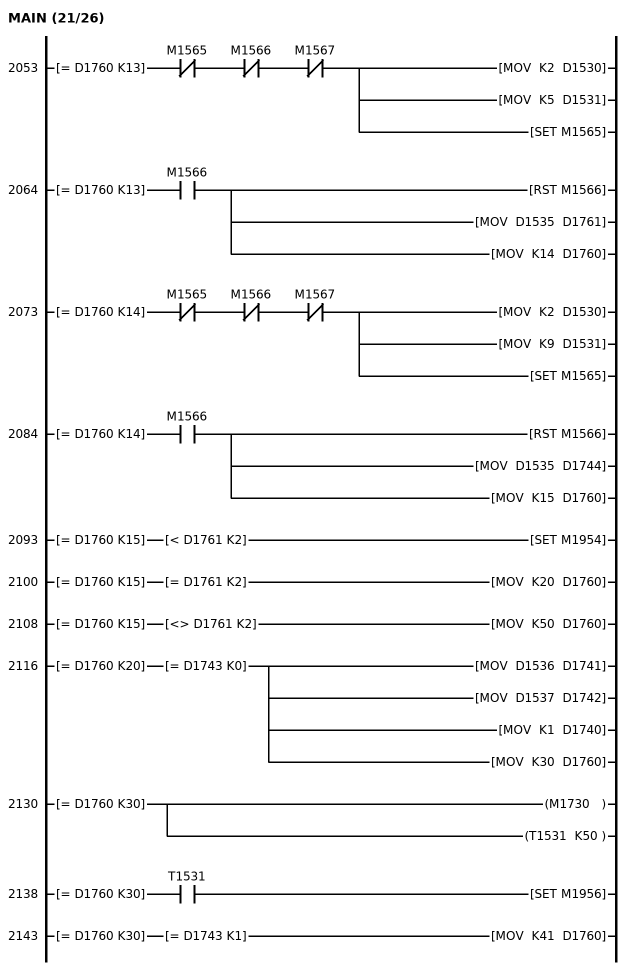
2053  LD=     D1760 K13
      ANI     M1565
      ANI     M1566
      ANI     M1567
      MOV     K2 D1530
      MOV     K5 D1531
      SET     M1565
2064  LD=     D1760 K13
      AND     M1566
      RST     M1566
      MOV     D1535 D1761
      MOV     K14 D1760
2073  LD=     D1760 K14
      ANI     M1565
      ANI     M1566
      ANI     M1567
      MOV     K2 D1530
      MOV     K9 D1531
      SET     M1565
2084  LD=     D1760 K14
      AND     M1566
      RST     M1566
      MOV     D1535 D1744
      MOV     K15 D1760
2093  LD=     D1760 K15
      AND<    D1761 K2
      SET     M1954
2100  LD=     D1760 K15
      AND=    D1761 K2
      MOV     K20 D1760
2108  LD=     D1760 K15
      AND<>   D1761 K2
      MOV     K50 D1760
2116  LD=     D1760 K20
      AND=    D1743 K0
      MOV     D1536 D1741
      MOV     D1537 D1742
      MOV     K1 D1740
      MOV     K30 D1760
2130  LD=     D1760 K30
      OUT     M1730
      OUT     T1531 K50
2138  LD=     D1760 K30
      AND     T1531
      SET     M1956
2143  LD=     D1760 K30
      AND=    D1743 K1
      MOV     K41 D1760
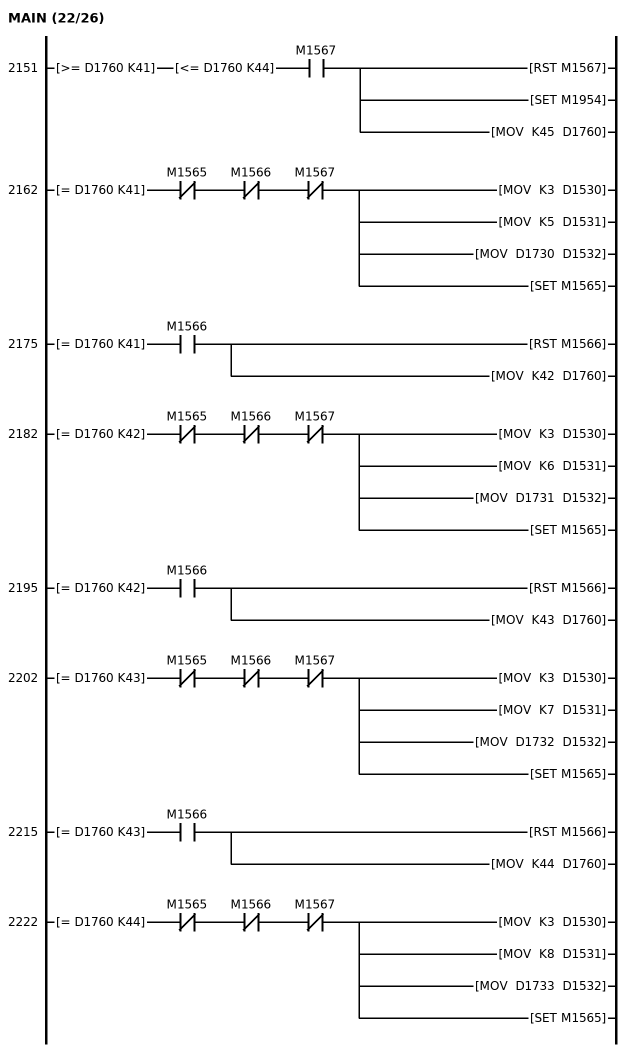
2151  LD>=    D1760 K41
      AND<=   D1760 K44
      AND     M1567
      RST     M1567
      SET     M1954
      MOV     K45 D1760
2162  LD=     D1760 K41
      ANI     M1565
      ANI     M1566
      ANI     M1567
      MOV     K3 D1530
      MOV     K5 D1531
      MOV     D1730 D1532
      SET     M1565
2175  LD=     D1760 K41
      AND     M1566
      RST     M1566
      MOV     K42 D1760
2182  LD=     D1760 K42
      ANI     M1565
      ANI     M1566
      ANI     M1567
      MOV     K3 D1530
      MOV     K6 D1531
      MOV     D1731 D1532
      SET     M1565
2195  LD=     D1760 K42
      AND     M1566
      RST     M1566
      MOV     K43 D1760
2202  LD=     D1760 K43
      ANI     M1565
      ANI     M1566
      ANI     M1567
      MOV     K3 D1530
      MOV     K7 D1531
      MOV     D1732 D1532
      SET     M1565
2215  LD=     D1760 K43
      AND     M1566
      RST     M1566
      MOV     K44 D1760
2222  LD=     D1760 K44
      ANI     M1565
      ANI     M1566
      ANI     M1567
      MOV     K3 D1530
      MOV     K8 D1531
      MOV     D1733 D1532
      SET     M1565
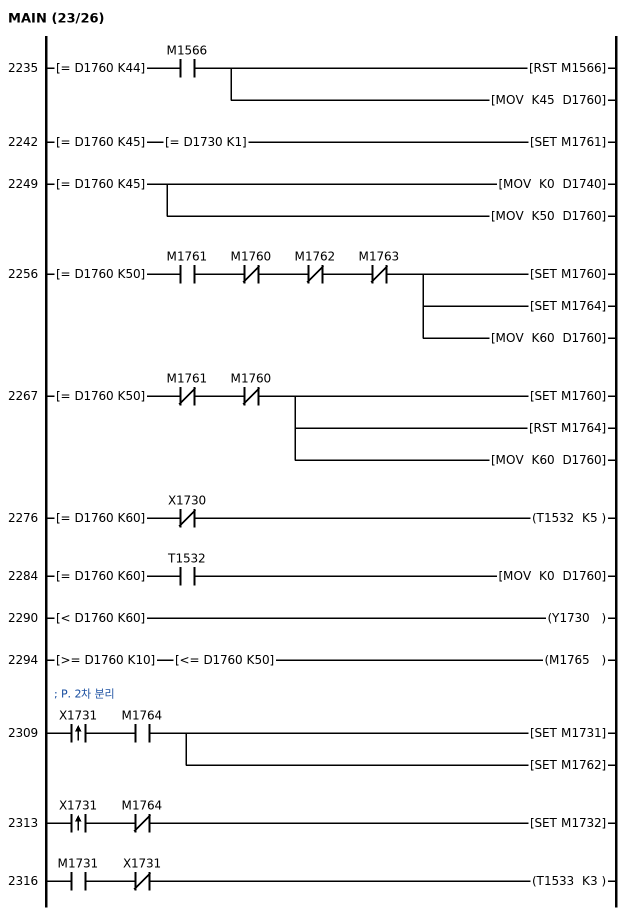
2235  LD=     D1760 K44
      AND     M1566
      RST     M1566
      MOV     K45 D1760
2242  LD=     D1760 K45
      AND=    D1730 K1
      SET     M1761
2249  LD=     D1760 K45
      MOV     K0 D1740
      MOV     K50 D1760
2256  LD=     D1760 K50
      AND     M1761
      ANI     M1760
      ANI     M1762
      ANI     M1763
      SET     M1760
      SET     M1764
      MOV     K60 D1760
2267  LD=     D1760 K50
      ANI     M1761
      ANI     M1760
      SET     M1760
      RST     M1764
      MOV     K60 D1760
2276  LD=     D1760 K60
      ANI     X1730
      OUT     T1532 K5
2284  LD=     D1760 K60
      AND     T1532
      MOV     K0 D1760
2290  LD<     D1760 K60
      OUT     Y1730
2294  LD>=    D1760 K10
      AND<=   D1760 K50
      OUT     M1765
; P. 2차 분리
2309  LDP     X1731
      AND     M1764
      SET     M1731
      SET     M1762
2313  LDP     X1731
      ANI     M1764
      SET     M1732
2316  LD      M1731
      ANI     X1731
      OUT     T1533 K3
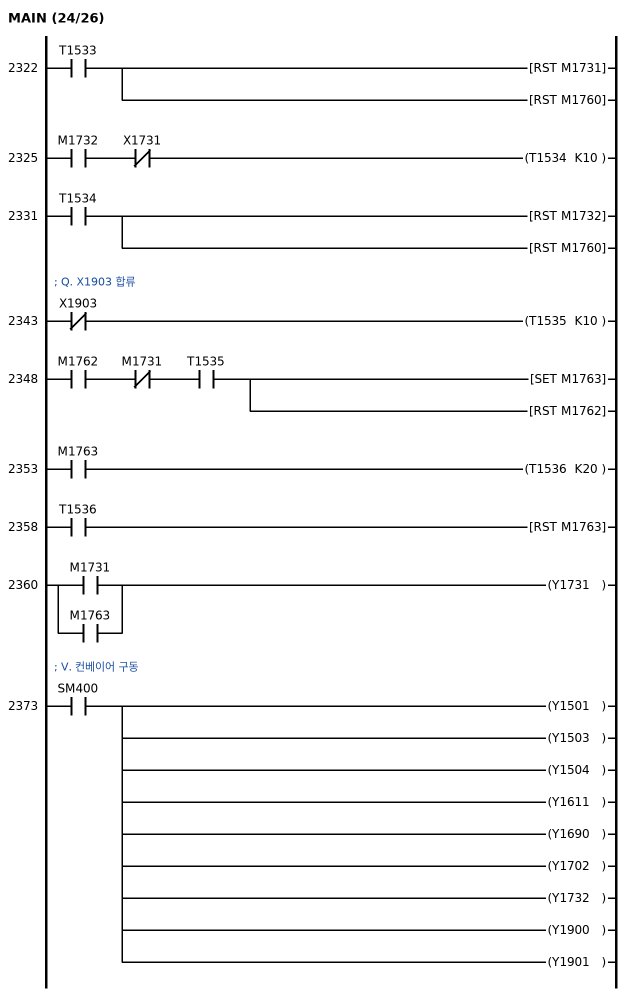
2322  LD      T1533
      RST     M1731
      RST     M1760
2325  LD      M1732
      ANI     X1731
      OUT     T1534 K10
2331  LD      T1534
      RST     M1732
      RST     M1760
; Q. X1903 합류
2343  LDI     X1903
      OUT     T1535 K10
2348  LD      M1762
      ANI     M1731
      AND     T1535
      SET     M1763
      RST     M1762
2353  LD      M1763
      OUT     T1536 K20
2358  LD      T1536
      RST     M1763
2360  LD      M1731
      OR      M1763
      OUT     Y1731
; V. 컨베이어 구동
2373  LD      SM400
      OUT     Y1501
      OUT     Y1503
      OUT     Y1504
      OUT     Y1611
      OUT     Y1690
      OUT     Y1702
      OUT     Y1732
      OUT     Y1900
      OUT     Y1901
